(* IEC 61131-3 sources: plc-iiot-stack/src/POUs/Json/FB_JsonFlatParser, 30 files *)

(* ---- FB_JsonFlatParser.decl.st ---- *)
// Назначение: разбор подмножества JSON для команд: один плоский объект, значения — строки (до
//             JSON_STR_LEN, escape-последовательности ASCII), числа по грамматике JSON (в диапазоне
//             REAL), true, false, null. Вложенные объекты и массивы, повторяющиеся ключи, лишние
//             символы после объекта — отказ с причиной eError и позицией uiErrorPos.
//             Порядок: Parse(sJson), затем GetString, GetNumber, FieldType по ключу.
// Автор:      kr0nsch
// Версия:     0.1.0
// Документ:   docs/plc_mqtt.md, раздел «Команды»
FUNCTION_BLOCK FB_JsonFlatParser
VAR_OUTPUT
    uiCount : UINT;                       // полей в разобранном объекте
    eError : E_JsonError := E_JsonError.None;
    uiErrorPos : UINT;                    // позиция ошибки (байт от 0)
END_VAR
VAR
    aFields : ARRAY[1..GVL_Const.JSON_MAX_FIELDS] OF ST_JsonField;
    uiPos : UINT;                         // текущая позиция разбора
    uiLen : UINT;                         // длина входа
    sTok : STRING(GVL_Const.JSON_STR_LEN);   // последний разобранный токен-строка (ключ или значение)
    lrTok : LREAL;                        // последнее разобранное число
    xTokInteger : BOOL;                   // число записано без дробной части и порядка
END_VAR

(* ---- Fail.method.decl.st ---- *)
// Зафиксировать ошибку разбора в текущей позиции; поля разобранного объекта сбрасываются.
METHOD PRIVATE Fail
VAR_INPUT
    eReason : E_JsonError;
END_VAR

(* ---- FieldIsInteger.method.decl.st ---- *)
// Поле sKey — число, записанное без дробной части и порядка (целое JSON Schema в строгом смысле).
METHOD FieldIsInteger : BOOL
VAR_INPUT
    sKey : STRING(GVL_Const.JSON_KEY_LEN);
END_VAR
VAR
    uiIdx : UINT;
END_VAR

(* ---- FieldIsInteger.method.impl.st ---- *)
uiIdx := FindField(sKey := sKey);
IF uiIdx > 0 THEN
    FieldIsInteger := aFields[uiIdx].eType = E_JsonType.Number AND aFields[uiIdx].xInteger;
END_IF

(* ---- FieldType.method.decl.st ---- *)
// Тип значения поля sKey; поля нет — Missing.
METHOD FieldType : E_JsonType
VAR_INPUT
    sKey : STRING(GVL_Const.JSON_KEY_LEN);
END_VAR
VAR
    uiIdx : UINT;
END_VAR

(* ---- FieldType.method.impl.st ---- *)
uiIdx := FindField(sKey := sKey);
IF uiIdx = 0 THEN
    FieldType := E_JsonType.Missing;
ELSE
    FieldType := aFields[uiIdx].eType;
END_IF

(* ---- FindField.method.decl.st ---- *)
// Индекс поля с ключом sKey (с учётом регистра); нет — 0.
METHOD FindField : UINT
VAR_INPUT
    sKey : STRING(GVL_Const.JSON_KEY_LEN);
END_VAR
VAR
    uiIdx : UINT;
END_VAR

(* ---- FindField.method.impl.st ---- *)
FindField := 0;
FOR uiIdx := 1 TO uiCount DO
    IF aFields[uiIdx].sKey = sKey THEN
        FindField := uiIdx;
        RETURN;
    END_IF
END_FOR

(* ---- GetBool.method.decl.st ---- *)
// Логическое значение поля sKey. TRUE — поле есть и это true или false; иначе xValue не меняется.
METHOD GetBool : BOOL
VAR_INPUT
    sKey : STRING(GVL_Const.JSON_KEY_LEN);
END_VAR
VAR_IN_OUT
    xValue : BOOL;
END_VAR
VAR
    uiIdx : UINT;
END_VAR

(* ---- GetBool.method.impl.st ---- *)
uiIdx := FindField(sKey := sKey);
IF uiIdx > 0 THEN
    IF aFields[uiIdx].eType = E_JsonType.Boolean THEN
        xValue := aFields[uiIdx].xBool;
        GetBool := TRUE;
    END_IF
END_IF

(* ---- GetNumber.method.decl.st ---- *)
// Числовое значение поля sKey. TRUE — поле есть и это число; иначе lrValue не меняется.
METHOD GetNumber : BOOL
VAR_INPUT
    sKey : STRING(GVL_Const.JSON_KEY_LEN);
END_VAR
VAR_IN_OUT
    lrValue : LREAL;
END_VAR
VAR
    uiIdx : UINT;
END_VAR

(* ---- GetNumber.method.impl.st ---- *)
uiIdx := FindField(sKey := sKey);
IF uiIdx > 0 THEN
    IF aFields[uiIdx].eType = E_JsonType.Number THEN
        lrValue := aFields[uiIdx].lrNumber;
        GetNumber := TRUE;
    END_IF
END_IF

(* ---- GetString.method.decl.st ---- *)
// Строковое значение поля sKey. TRUE — поле есть и это строка; иначе sValue не меняется.
METHOD GetString : BOOL
VAR_INPUT
    sKey : STRING(GVL_Const.JSON_KEY_LEN);
END_VAR
VAR_IN_OUT
    sValue : STRING(GVL_Const.JSON_STR_LEN);
END_VAR
VAR
    uiIdx : UINT;
END_VAR

(* ---- GetString.method.impl.st ---- *)
uiIdx := FindField(sKey := sKey);
IF uiIdx > 0 THEN
    IF aFields[uiIdx].eType = E_JsonType.Text THEN
        sValue := aFields[uiIdx].sText;
        GetString := TRUE;
    END_IF
END_IF

(* ---- HexValue.method.decl.st ---- *)
// Значение шестнадцатеричной цифры 0..15; не цифра — -1.
METHOD PRIVATE HexValue : INT
VAR_INPUT
    bDigit : BYTE;
END_VAR

(* ---- HexValue.method.impl.st ---- *)
IF bDigit >= GVL_Const.ASCII_ZERO AND bDigit <= GVL_Const.ASCII_NINE THEN
    HexValue := BYTE_TO_INT(bDigit - GVL_Const.ASCII_ZERO);
ELSIF bDigit >= GVL_Const.ASCII_LOWER_A AND bDigit <= GVL_Const.ASCII_LOWER_F THEN
    HexValue := BYTE_TO_INT(bDigit - GVL_Const.ASCII_LOWER_A + GVL_Const.HEX_LETTER_START);
ELSIF bDigit >= GVL_Const.ASCII_UPPER_A AND bDigit <= GVL_Const.ASCII_UPPER_F THEN
    HexValue := BYTE_TO_INT(bDigit - GVL_Const.ASCII_UPPER_A + GVL_Const.HEX_LETTER_START);
ELSE
    HexValue := -1;
END_IF

(* ---- KeyAt.method.decl.st ---- *)
// Ключ поля с номером uiIdx (1..uiCount); вне диапазона — пустая строка.
METHOD KeyAt : STRING(GVL_Const.JSON_KEY_LEN)
VAR_INPUT
    uiIdx : UINT;
END_VAR

(* ---- KeyAt.method.impl.st ---- *)
IF uiIdx >= 1 AND uiIdx <= uiCount THEN
    KeyAt := aFields[uiIdx].sKey;
END_IF

(* ---- MatchLiteral.method.decl.st ---- *)
// Сравнить вход с литералом (true, false, null) и сдвинуть позицию за него. FALSE — ошибка Syntax.
METHOD PRIVATE MatchLiteral : BOOL
VAR_IN_OUT CONSTANT
    // lint:allow STL007 параметр VAR_IN_OUT CONSTANT — ссылка только для чтения, а не константа
    sJson : STRING(GVL_Const.MQTT_CMD_PAYLOAD_LEN);
END_VAR
VAR_INPUT
    sLiteral : STRING(GVL_Const.JSON_LITERAL_LEN);
END_VAR
VAR
    uiLitLen : UINT;
    uiIdx : UINT;
END_VAR

(* ---- MatchLiteral.method.impl.st ---- *)
uiLitLen := INT_TO_UINT(LEN(sLiteral));
IF uiPos + uiLitLen > uiLen THEN
    Fail(eReason := E_JsonError.Syntax);
    RETURN;
END_IF
FOR uiIdx := 0 TO uiLitLen - 1 DO
    IF sJson[uiPos + uiIdx] <> sLiteral[uiIdx] THEN
        uiPos := uiPos + uiIdx;
        Fail(eReason := E_JsonError.Syntax);
        RETURN;
    END_IF
END_FOR
uiPos := uiPos + uiLitLen;
MatchLiteral := TRUE;

(* ---- Parse.method.decl.st ---- *)
// Разобрать объект. TRUE — разбор успешен (uiCount полей); FALSE — eError и uiErrorPos.
METHOD Parse : BOOL
VAR_IN_OUT CONSTANT
    // lint:allow STL007 параметр VAR_IN_OUT CONSTANT — ссылка только для чтения, а не константа
    sJson : STRING(GVL_Const.MQTT_CMD_PAYLOAD_LEN);
END_VAR
VAR
    bCh : BYTE;
    stField : ST_JsonField;
END_VAR

(* ---- Parse.method.impl.st ---- *)
uiCount := 0;
eError := E_JsonError.None;
uiErrorPos := 0;
uiPos := 0;
uiLen := 0;
WHILE uiLen < GVL_Const.MQTT_CMD_PAYLOAD_LEN AND_THEN sJson[uiLen] <> GVL_Const.ASCII_NUL DO
    uiLen := uiLen + 1;
END_WHILE

SkipSpace(sJson := sJson);
IF uiPos >= uiLen THEN
    Fail(eReason := E_JsonError.Empty);
    RETURN;
END_IF
IF Peek(sJson := sJson) <> GVL_Const.ASCII_LBRACE THEN
    Fail(eReason := E_JsonError.Syntax);
    RETURN;
END_IF
uiPos := uiPos + 1;
SkipSpace(sJson := sJson);

IF Peek(sJson := sJson) = GVL_Const.ASCII_RBRACE THEN
    uiPos := uiPos + 1;      // пустой объект {}
ELSE
    WHILE TRUE DO
        // ключ
        IF Peek(sJson := sJson) <> GVL_Const.ASCII_QUOTE THEN
            Fail(eReason := E_JsonError.Syntax);
            RETURN;
        END_IF
        IF NOT ParseText(sJson := sJson, uiMaxLen := GVL_Const.JSON_KEY_LEN, eTooLong := E_JsonError.KeyTooLong) THEN
            RETURN;
        END_IF
        stField.sKey := sTok;
        stField.sText := '';
        stField.lrNumber := 0.0;
        stField.xInteger := FALSE;
        stField.xBool := FALSE;
        SkipSpace(sJson := sJson);
        IF Peek(sJson := sJson) <> GVL_Const.ASCII_COLON THEN
            Fail(eReason := E_JsonError.Syntax);
            RETURN;
        END_IF
        uiPos := uiPos + 1;
        SkipSpace(sJson := sJson);

        // значение
        bCh := Peek(sJson := sJson);
        IF bCh = GVL_Const.ASCII_QUOTE THEN
            IF NOT ParseText(sJson := sJson, uiMaxLen := GVL_Const.JSON_STR_LEN,
                             eTooLong := E_JsonError.ValueTooLong) THEN
                RETURN;
            END_IF
            stField.eType := E_JsonType.Text;
            stField.sText := sTok;
        ELSIF bCh = GVL_Const.ASCII_MINUS OR (bCh >= GVL_Const.ASCII_ZERO AND bCh <= GVL_Const.ASCII_NINE) THEN
            IF NOT ParseNumber(sJson := sJson) THEN
                RETURN;
            END_IF
            stField.eType := E_JsonType.Number;
            stField.lrNumber := lrTok;
            stField.xInteger := xTokInteger;
        ELSIF bCh = GVL_Const.ASCII_LOWER_T THEN
            IF NOT MatchLiteral(sJson := sJson, sLiteral := 'true') THEN
                RETURN;
            END_IF
            stField.eType := E_JsonType.Boolean;
            stField.xBool := TRUE;
        ELSIF bCh = GVL_Const.ASCII_LOWER_F THEN
            IF NOT MatchLiteral(sJson := sJson, sLiteral := 'false') THEN
                RETURN;
            END_IF
            stField.eType := E_JsonType.Boolean;
        ELSIF bCh = GVL_Const.ASCII_LOWER_N THEN
            IF NOT MatchLiteral(sJson := sJson, sLiteral := 'null') THEN
                RETURN;
            END_IF
            stField.eType := E_JsonType.NullValue;
        ELSIF bCh = GVL_Const.ASCII_LBRACE OR bCh = GVL_Const.ASCII_LBRACKET THEN
            Fail(eReason := E_JsonError.Nested);
            RETURN;
        ELSE
            Fail(eReason := E_JsonError.Syntax);
            RETURN;
        END_IF

        IF FindField(sKey := stField.sKey) > 0 THEN
            Fail(eReason := E_JsonError.Duplicate);
            RETURN;
        END_IF
        IF uiCount >= GVL_Const.JSON_MAX_FIELDS THEN
            Fail(eReason := E_JsonError.TooManyFields);
            RETURN;
        END_IF
        uiCount := uiCount + 1;
        aFields[uiCount] := stField;

        SkipSpace(sJson := sJson);
        bCh := Peek(sJson := sJson);
        IF bCh = GVL_Const.ASCII_COMMA THEN
            uiPos := uiPos + 1;
            SkipSpace(sJson := sJson);
        ELSIF bCh = GVL_Const.ASCII_RBRACE THEN
            uiPos := uiPos + 1;
            EXIT;
        ELSE
            Fail(eReason := E_JsonError.Syntax);
            RETURN;
        END_IF
    END_WHILE
END_IF

SkipSpace(sJson := sJson);
IF uiPos < uiLen THEN
    Fail(eReason := E_JsonError.Trailing);
    RETURN;
END_IF
Parse := TRUE;

(* ---- ParseNumber.method.decl.st ---- *)
// Разобрать число по грамматике JSON -?(0|[1-9]d*)(.d+)?([eE][+-]?d+)? в lrTok. Нарушение грамматики,
// больше JSON_MANTISSA_DIGITS_MAX цифр, больше JSON_EXP_DIGITS_MAX цифр порядка, |x| > REAL_ABS_MAX —
// ошибка BadNumber.
METHOD PRIVATE ParseNumber : BOOL
VAR_IN_OUT CONSTANT
    // lint:allow STL007 параметр VAR_IN_OUT CONSTANT — ссылка только для чтения, а не константа
    sJson : STRING(GVL_Const.MQTT_CMD_PAYLOAD_LEN);
END_VAR
VAR
    bCh : BYTE;
    xNegative : BOOL;
    xExpNegative : BOOL;
    lrMantissa : LREAL;
    uiDigits : UINT;       // цифр мантиссы
    iFracDigits : INT;     // цифр после точки
    uiExpDigits : UINT;
    iExp : INT;
    xHasExp : BOOL;
END_VAR

(* ---- ParseNumber.method.impl.st ---- *)
lrTok := 0.0;
xTokInteger := FALSE;
IF Peek(sJson := sJson) = GVL_Const.ASCII_MINUS THEN
    xNegative := TRUE;
    uiPos := uiPos + 1;
END_IF
bCh := Peek(sJson := sJson);
IF bCh < GVL_Const.ASCII_ZERO OR bCh > GVL_Const.ASCII_NINE THEN
    Fail(eReason := E_JsonError.BadNumber);
    RETURN;
END_IF

// целая часть: 0 или цифры без ведущего нуля
IF bCh = GVL_Const.ASCII_ZERO THEN
    uiPos := uiPos + 1;
    uiDigits := 1;
    bCh := Peek(sJson := sJson);
    IF bCh >= GVL_Const.ASCII_ZERO AND bCh <= GVL_Const.ASCII_NINE THEN
        Fail(eReason := E_JsonError.BadNumber);
        RETURN;
    END_IF
ELSE
    WHILE bCh >= GVL_Const.ASCII_ZERO AND bCh <= GVL_Const.ASCII_NINE DO
        lrMantissa := lrMantissa * ULINT_TO_LREAL(GVL_Const.DECIMAL_BASE) + BYTE_TO_LREAL(bCh - GVL_Const.ASCII_ZERO);
        uiDigits := uiDigits + 1;
        uiPos := uiPos + 1;
        bCh := Peek(sJson := sJson);
    END_WHILE
END_IF

// дробная часть
IF bCh = GVL_Const.ASCII_DOT THEN
    uiPos := uiPos + 1;
    bCh := Peek(sJson := sJson);
    IF bCh < GVL_Const.ASCII_ZERO OR bCh > GVL_Const.ASCII_NINE THEN
        Fail(eReason := E_JsonError.BadNumber);
        RETURN;
    END_IF
    WHILE bCh >= GVL_Const.ASCII_ZERO AND bCh <= GVL_Const.ASCII_NINE DO
        lrMantissa := lrMantissa * ULINT_TO_LREAL(GVL_Const.DECIMAL_BASE) + BYTE_TO_LREAL(bCh - GVL_Const.ASCII_ZERO);
        uiDigits := uiDigits + 1;
        iFracDigits := iFracDigits + 1;
        uiPos := uiPos + 1;
        bCh := Peek(sJson := sJson);
    END_WHILE
END_IF
IF uiDigits > GVL_Const.JSON_MANTISSA_DIGITS_MAX THEN
    Fail(eReason := E_JsonError.BadNumber);
    RETURN;
END_IF

// порядок
IF bCh = GVL_Const.ASCII_LOWER_E OR bCh = GVL_Const.ASCII_UPPER_E THEN
    xHasExp := TRUE;
    uiPos := uiPos + 1;
    bCh := Peek(sJson := sJson);
    IF bCh = GVL_Const.ASCII_MINUS THEN
        xExpNegative := TRUE;
        uiPos := uiPos + 1;
    ELSIF bCh = GVL_Const.ASCII_PLUS THEN
        uiPos := uiPos + 1;
    END_IF
    bCh := Peek(sJson := sJson);
    IF bCh < GVL_Const.ASCII_ZERO OR bCh > GVL_Const.ASCII_NINE THEN
        Fail(eReason := E_JsonError.BadNumber);
        RETURN;
    END_IF
    WHILE bCh >= GVL_Const.ASCII_ZERO AND bCh <= GVL_Const.ASCII_NINE DO
        IF uiExpDigits >= GVL_Const.JSON_EXP_DIGITS_MAX THEN
            Fail(eReason := E_JsonError.BadNumber);
            RETURN;
        END_IF
        iExp := iExp * ULINT_TO_INT(GVL_Const.DECIMAL_BASE) + BYTE_TO_INT(bCh - GVL_Const.ASCII_ZERO);
        uiExpDigits := uiExpDigits + 1;
        uiPos := uiPos + 1;
        bCh := Peek(sJson := sJson);
    END_WHILE
    IF xExpNegative THEN
        iExp := -iExp;
    END_IF
END_IF

lrTok := lrMantissa * EXPT(ULINT_TO_LREAL(GVL_Const.DECIMAL_BASE), INT_TO_LREAL(iExp - iFracDigits));
xTokInteger := iFracDigits = 0 AND NOT xHasExp;
IF xNegative THEN
    lrTok := -lrTok;
END_IF
IF NOT (ABS(lrTok) <= GVL_Const.REAL_ABS_MAX) THEN
    Fail(eReason := E_JsonError.BadNumber);
    RETURN;
END_IF
ParseNumber := TRUE;

(* ---- ParseText.method.decl.st ---- *)
// Разобрать строку в кавычках (позиция — на открывающей кавычке) в sTok. Длиннее uiMaxLen — ошибка
// eTooLong. Управляющие символы без экранирования, незакрытая строка — Syntax; \u вне ASCII — BadEscape.
METHOD PRIVATE ParseText : BOOL
VAR_IN_OUT CONSTANT
    // lint:allow STL007 параметр VAR_IN_OUT CONSTANT — ссылка только для чтения, а не константа
    sJson : STRING(GVL_Const.MQTT_CMD_PAYLOAD_LEN);
END_VAR
VAR_INPUT
    uiMaxLen : UINT;
    eTooLong : E_JsonError;
END_VAR
VAR
    bCh : BYTE;
    uiOut : UINT;          // длина sTok
    uiHex : UINT;
    iDigit : INT;
    uiCode : UINT;         // код символа \uXXXX
END_VAR

(* ---- ParseText.method.impl.st ---- *)
sTok := '';
uiOut := 0;
uiPos := uiPos + 1;   // за открывающую кавычку
WHILE TRUE DO
    IF uiPos >= uiLen THEN
        Fail(eReason := E_JsonError.Syntax);   // строка не закрыта
        RETURN;
    END_IF
    bCh := sJson[uiPos];
    IF bCh = GVL_Const.ASCII_QUOTE THEN
        uiPos := uiPos + 1;
        EXIT;
    END_IF
    IF bCh <= GVL_Const.ASCII_CTRL_LAST THEN
        Fail(eReason := E_JsonError.Syntax);
        RETURN;
    END_IF
    IF bCh = GVL_Const.ASCII_BACKSLASH THEN
        uiPos := uiPos + 1;
        IF uiPos >= uiLen THEN
            Fail(eReason := E_JsonError.Syntax);
            RETURN;
        END_IF
        bCh := sJson[uiPos];
        // после обратной косой черты: кавычка, обратная и прямая косая черта дают сами себя
        IF bCh = GVL_Const.ASCII_LOWER_N THEN
            bCh := GVL_Const.ASCII_LF;
        ELSIF bCh = GVL_Const.ASCII_LOWER_R THEN
            bCh := GVL_Const.ASCII_CR;
        ELSIF bCh = GVL_Const.ASCII_LOWER_T THEN
            bCh := GVL_Const.ASCII_TAB;
        ELSIF bCh = GVL_Const.ASCII_LOWER_B THEN
            bCh := GVL_Const.ASCII_BS;
        ELSIF bCh = GVL_Const.ASCII_LOWER_F THEN
            bCh := GVL_Const.ASCII_FF;
        ELSIF bCh = GVL_Const.ASCII_LOWER_U THEN
            uiCode := 0;
            FOR uiHex := 1 TO GVL_Const.HEX_DIGITS_ESCAPE DO
                IF uiPos + uiHex >= uiLen THEN
                    Fail(eReason := E_JsonError.BadEscape);
                    RETURN;
                END_IF
                iDigit := HexValue(bDigit := sJson[uiPos + uiHex]);
                IF iDigit < 0 THEN
                    Fail(eReason := E_JsonError.BadEscape);
                    RETURN;
                END_IF
                uiCode := uiCode * GVL_Const.HEX_BASE + INT_TO_UINT(iDigit);
            END_FOR
            // поддерживаются только символы ASCII без нуля
            IF uiCode = 0 OR uiCode > BYTE_TO_UINT(GVL_Const.ASCII_LAST) THEN
                Fail(eReason := E_JsonError.BadEscape);
                RETURN;
            END_IF
            uiPos := uiPos + GVL_Const.HEX_DIGITS_ESCAPE;
            bCh := UINT_TO_BYTE(uiCode);
        ELSIF bCh <> GVL_Const.ASCII_QUOTE AND bCh <> GVL_Const.ASCII_BACKSLASH AND bCh <> GVL_Const.ASCII_SLASH THEN
            Fail(eReason := E_JsonError.BadEscape);
            RETURN;
        END_IF
    END_IF
    IF uiOut >= uiMaxLen THEN
        Fail(eReason := eTooLong);
        RETURN;
    END_IF
    sTok[uiOut] := bCh;
    uiOut := uiOut + 1;
    sTok[uiOut] := GVL_Const.ASCII_NUL;
    uiPos := uiPos + 1;
END_WHILE
ParseText := TRUE;

(* ---- Peek.method.decl.st ---- *)
// Текущий байт входа; за концом — 0.
METHOD PRIVATE Peek : BYTE
VAR_IN_OUT CONSTANT
    // lint:allow STL007 параметр VAR_IN_OUT CONSTANT — ссылка только для чтения, а не константа
    sJson : STRING(GVL_Const.MQTT_CMD_PAYLOAD_LEN);
END_VAR

(* ---- Peek.method.impl.st ---- *)
IF uiPos < uiLen THEN
    Peek := sJson[uiPos];
ELSE
    Peek := GVL_Const.ASCII_NUL;
END_IF

(* ---- SkipSpace.method.decl.st ---- *)
// Пропустить пробельные символы JSON: пробел, табуляция, перевод строки, возврат каретки.
METHOD PRIVATE SkipSpace
VAR_IN_OUT CONSTANT
    // lint:allow STL007 параметр VAR_IN_OUT CONSTANT — ссылка только для чтения, а не константа
    sJson : STRING(GVL_Const.MQTT_CMD_PAYLOAD_LEN);
END_VAR
VAR
    bCh : BYTE;
END_VAR

(* ---- SkipSpace.method.impl.st ---- *)
WHILE uiPos < uiLen DO
    bCh := sJson[uiPos];
    IF bCh = GVL_Const.ASCII_SPACE OR bCh = GVL_Const.ASCII_TAB OR bCh = GVL_Const.ASCII_LF
       OR bCh = GVL_Const.ASCII_CR THEN
        uiPos := uiPos + 1;
    ELSE
        EXIT;
    END_IF
END_WHILE
